// Stato di una valvola per l'HMI.
TYPE ST_HmiValveSts :
STRUCT
	bSet			: BOOL;		// uscita "set"
	bReset			: BOOL;		// uscita "reset" (bistabile)
	bFbSet			: BOOL;		// conferma lato set
	bFbReset		: BOOL;		// conferma lato reset
END_STRUCT
END_TYPE

(* stored: Version 1.1.0.1, ProductVersion 3.1.4024.12
   DUT ST_HmiValveSts: Id {aee226ff-34f4-4dec-a92e-413badc6ba1d} *)
